TYPE typeMessage :
STRUCT
	//defines a list of messages to display for each type of message
	
	message: ARRAY [0..GlobalMessages.gNumMessagesPerType] OF BOOL; //TRUE if the message is active to be written to the message box	
	text:ARRAY[0..GlobalMessages.gNumMessagesPerType] OF STRING(255); //the text of each message to be written
	messageActive: ARRAY [0..GlobalMessages.gNumMessagesPerType] OF BOOL; //TRUE if the message has been written to the message box
	messageTimeActive: ARRAY [0..GlobalMessages.gNumMessagesPerType] OF UDINT; //scan time occurrence of each message to compare
	
	topMessage:STRING(255); //top message to display
	
	allMessage:STRING;
	
END_STRUCT
END_TYPE

(* stored: Version 1.1.0.1, ProductVersion 3.1.4024.12
   DUT typeMessage: Id {221336c1-ab93-4c6c-ba86-6e53bedca566} *)
